PROGRAM PRG_StationProcessSettings
VAR
    bInitialised : BOOL;
    bWritePending : BOOL;
    bWriteStart : BOOL;
    bWriteBusySeen : BOOL;
    fbWritePersistentData : FB_WritePersistentData;
    stDefaultPatch : ST_PatchProcessSettings;
    stDefaultVision : ST_CameraProcessSettings;
    bSafetySaveAcceptedPending : BOOL;
    bSafetySettingsInitialised : BOOL;
    bVisionPbupSavePending : BOOL;
    bVisionPbupSaveInFlight : BOOL;
END_VAR

IF NOT bInitialised THEN
    // Preserve retained values; new speeds and delay are applied through Patch Settings.
    IF NOT ((GVL_Persistent.stPatchProcessSettings.lrDriveMotorVelocity >= 0.1) AND (GVL_Persistent.stPatchProcessSettings.lrDriveMotorVelocity <= 40)
        AND (GVL_Persistent.stPatchProcessSettings.lrPatchFeedRollVelocity >= 0.1) AND (GVL_Persistent.stPatchProcessSettings.lrPatchFeedRollVelocity <= 200)
        AND (GVL_Persistent.stPatchProcessSettings.lrWasteRollVelocity >= 0.1) AND (GVL_Persistent.stPatchProcessSettings.lrWasteRollVelocity <= 50)
        AND (GVL_Persistent.stPatchProcessSettings.udiReleaseMs >= 100) AND (GVL_Persistent.stPatchProcessSettings.udiReleaseMs <= 15000)
        AND (GVL_Persistent.stPatchProcessSettings.udiAirBlowDelayMs >= 0) AND (GVL_Persistent.stPatchProcessSettings.udiAirBlowDelayMs <= 5000)
        AND (GVL_Persistent.stPatchProcessSettings.udiDriveStopDelayMs >= 0) AND (GVL_Persistent.stPatchProcessSettings.udiDriveStopDelayMs <= 5000)) THEN
        GVL_Persistent.stPatchProcessSettings := stDefaultPatch;
        GVL_HMI.sPatchSettingsMessage := 'Stored values invalid: defaults loaded. Review and Apply.';
    ELSE
        GVL_HMI.sPatchSettingsMessage := 'Ready';
    END_IF
    GVL_HMI.stPatchProcessEdit := GVL_Persistent.stPatchProcessSettings;
    IF NOT ((GVL_Persistent.stVisionProcessSettings.udiMovingTriggerDelayMs >= 0) AND (GVL_Persistent.stVisionProcessSettings.udiMovingTriggerDelayMs <= 1000)
        AND (GVL_Persistent.stVisionProcessSettings.udiRotaryConfirmMs >= 1000) AND (GVL_Persistent.stVisionProcessSettings.udiRotaryConfirmMs <= 3000)) THEN
        GVL_Persistent.stVisionProcessSettings := stDefaultVision;
        GVL_HMI.sVisionSettingsMessage := 'Stored values invalid: defaults loaded. Review and Apply.';
    ELSE
        GVL_HMI.sVisionSettingsMessage := 'Ready';
    END_IF
    GVL_HMI.stVisionProcessEdit := GVL_Persistent.stVisionProcessSettings;
    bInitialised := TRUE;
END_IF

// Initialize the new boundary independently, including after an online source change.
IF NOT bSafetySettingsInitialised THEN
    // Reuse the existing retained door threshold; do not reset other process settings.
    IF NOT ((GVL_Config.rMainDoorHotTemperatureLimitC >= 20.0)
        AND (GVL_Config.rMainDoorHotTemperatureLimitC <= 40.0)) THEN
        GVL_Config.rMainDoorHotTemperatureLimitC := 40.0;
        GVL_HMI.sSafetySettingsMessage := 'Stored limit invalid: 40 C loaded. Review and Apply.';
    ELSE
        GVL_HMI.sSafetySettingsMessage := 'Ready';
    END_IF
    GVL_HMI.rSafetyDoorHotLimitEditC := GVL_Config.rMainDoorHotTemperatureLimitC;
    bSafetySettingsInitialised := TRUE;
END_IF

// Use existing machine status; apply before PRG_Main starts any new process.
GVL_HMI.bStationSettingsAllowed :=
    ((GVL_MASTER.stStatus.eMachineState = E_MachineState.Stopped)
     OR (GVL_MASTER.stStatus.eMachineState = E_MachineState.ReadyToStart))
    AND NOT GVL_MASTER.stStatus.stPatchDispense.bBusy
    AND NOT GVL_MASTER.stStatus.stHeatStake.bBusy
    AND NOT GVL_MASTER.stStatus.stVision.bBusy
    AND NOT GVL_Motion.stPatchFeedStatus.bBusy
    AND NOT GVL_Motion.stPatchFeedStatus.bDriveBusy
    AND NOT GVL_Motion.AxisDriveMotor.bMoving
    AND NOT GVL_Motion.AxisPatchFeedRollMotor.bMoving
    AND NOT GVL_Motion.AxisWasteRollMotor.bMoving;
bWriteStart := FALSE;

// Cancel wins over Apply. Consume command BOOLs so the HMI can issue another request.
IF GVL_HMI.bPatchSettingsCancel THEN
    GVL_HMI.stPatchProcessEdit := GVL_Persistent.stPatchProcessSettings;
    GVL_HMI.sPatchSettingsMessage := 'Edits cancelled';
ELSIF GVL_HMI.bPatchSettingsApply THEN
    IF NOT GVL_HMI.bStationSettingsAllowed THEN
        GVL_HMI.sPatchSettingsMessage := 'Apply rejected: stop machine and motion first';
    ELSIF GVL_HMI.bStationSettingsSaving THEN
        GVL_HMI.sPatchSettingsMessage := 'Apply rejected: save in progress';
    ELSIF NOT ((GVL_HMI.stPatchProcessEdit.lrDriveMotorVelocity >= 0.1) AND (GVL_HMI.stPatchProcessEdit.lrDriveMotorVelocity <= 40)
        AND (GVL_HMI.stPatchProcessEdit.lrPatchFeedRollVelocity >= 0.1) AND (GVL_HMI.stPatchProcessEdit.lrPatchFeedRollVelocity <= 200)
        AND (GVL_HMI.stPatchProcessEdit.lrWasteRollVelocity >= 0.1) AND (GVL_HMI.stPatchProcessEdit.lrWasteRollVelocity <= 50)
        AND (GVL_HMI.stPatchProcessEdit.udiReleaseMs >= 100) AND (GVL_HMI.stPatchProcessEdit.udiReleaseMs <= 15000)
        AND (GVL_HMI.stPatchProcessEdit.udiAirBlowDelayMs >= 0) AND (GVL_HMI.stPatchProcessEdit.udiAirBlowDelayMs <= 5000)
        AND (GVL_HMI.stPatchProcessEdit.udiDriveStopDelayMs >= 0) AND (GVL_HMI.stPatchProcessEdit.udiDriveStopDelayMs <= 5000)) THEN
        GVL_HMI.sPatchSettingsMessage := 'Apply rejected: value outside allowed range';
    ELSE
        GVL_Persistent.stPatchProcessSettings := GVL_HMI.stPatchProcessEdit;
        bWritePending := TRUE;
        GVL_HMI.bStationSettingsSaveError := FALSE;
        GVL_HMI.udiStationSettingsSaveErrorId := 0;
        GVL_HMI.sPatchSettingsMessage := 'Applied - saving';
    END_IF
END_IF
GVL_HMI.bPatchSettingsApply := FALSE;
GVL_HMI.bPatchSettingsCancel := FALSE;
GVL_HMI.stPatchProcessApplied := GVL_Persistent.stPatchProcessSettings;

// Cancel wins over Apply. Consume command BOOLs so the HMI can issue another request.
IF GVL_HMI.bVisionSettingsCancel THEN
    GVL_HMI.stVisionProcessEdit := GVL_Persistent.stVisionProcessSettings;
    GVL_HMI.sVisionSettingsMessage := 'Edits cancelled';
ELSIF GVL_HMI.bVisionSettingsApply THEN
    IF NOT GVL_HMI.bStationSettingsAllowed THEN
        GVL_HMI.sVisionSettingsMessage := 'Apply rejected: stop machine and motion first';
    ELSIF GVL_HMI.bStationSettingsSaving THEN
        GVL_HMI.sVisionSettingsMessage := 'Apply rejected: save in progress';
    ELSIF NOT ((GVL_HMI.stVisionProcessEdit.udiMovingTriggerDelayMs >= 0) AND (GVL_HMI.stVisionProcessEdit.udiMovingTriggerDelayMs <= 1000)
        AND (GVL_HMI.stVisionProcessEdit.udiRotaryConfirmMs >= 1000) AND (GVL_HMI.stVisionProcessEdit.udiRotaryConfirmMs <= 3000)) THEN
        GVL_HMI.sVisionSettingsMessage := 'Apply rejected: value outside allowed range';
    ELSE
        GVL_Persistent.stVisionProcessSettings := GVL_HMI.stVisionProcessEdit;
        bWritePending := TRUE;
        GVL_HMI.bStationSettingsSaveError := FALSE;
        GVL_HMI.udiStationSettingsSaveErrorId := 0;
        GVL_HMI.sVisionSettingsMessage := 'Applied - saving';
    END_IF
END_IF
GVL_HMI.bVisionSettingsApply := FALSE;
GVL_HMI.bVisionSettingsCancel := FALSE;
GVL_HMI.stVisionProcessApplied := GVL_Persistent.stVisionProcessSettings;

// Safety settings are accepted only while Stopped and all existing settings/motion gates are clear.
GVL_HMI.bSafetySettingsAllowed := GVL_HMI.bStationSettingsAllowed
    AND (GVL_MASTER.stStatus.eMachineState = E_MachineState.Stopped)
    AND NOT GVL_MASTER.stCommand.bReset;
IF GVL_HMI.bSafetySettingsCancel THEN
    GVL_HMI.rSafetyDoorHotLimitEditC := GVL_Config.rMainDoorHotTemperatureLimitC;
    GVL_HMI.sSafetySettingsMessage := 'Edits cancelled';
ELSIF GVL_HMI.bSafetySettingsApply THEN
    IF NOT GVL_HMI.bSafetySettingsAllowed THEN
        GVL_HMI.sSafetySettingsMessage := 'Apply rejected: machine must be Stopped and idle';
    ELSIF GVL_HMI.bStationSettingsSaving THEN
        GVL_HMI.sSafetySettingsMessage := 'Apply rejected: save in progress';
    ELSIF NOT ((GVL_HMI.rSafetyDoorHotLimitEditC >= 20.0)
        AND (GVL_HMI.rSafetyDoorHotLimitEditC <= 40.0)) THEN
        GVL_HMI.sSafetySettingsMessage := 'Apply rejected: allowed range 20 to 40 C';
    ELSE
        GVL_Config.rMainDoorHotTemperatureLimitC := GVL_HMI.rSafetyDoorHotLimitEditC;
        bWritePending := TRUE;
        bSafetySaveAcceptedPending := TRUE;
        GVL_HMI.bStationSettingsSaveError := FALSE;
        GVL_HMI.udiStationSettingsSaveErrorId := 0;
        GVL_HMI.sSafetySettingsMessage := 'Applied - saving';
    END_IF
END_IF
GVL_HMI.bSafetySettingsApply := FALSE;
GVL_HMI.bSafetySettingsCancel := FALSE;
GVL_HMI.rSafetyDoorHotLimitAppliedC := GVL_Config.rMainDoorHotTemperatureLimitC;

// Request is latched by PRG_Main after this program; consume it on the next scan.
IF GVL_HMI.bVisionPbupSaveRequest THEN
    GVL_HMI.bVisionPbupSaveRequest := FALSE;
    bWritePending := TRUE;
    bVisionPbupSavePending := TRUE;
    GVL_HMI.bVisionPbupSaveError := FALSE;
    GVL_HMI.udiVisionPbupSaveErrorId := 0;
    GVL_HMI.sVisionPbupSaveStatus := 'PBUP state: save pending';
END_IF
IF bWritePending AND NOT fbWritePersistentData.BUSY THEN
    bWriteStart := TRUE;
    bWritePending := FALSE;
    bWriteBusySeen := FALSE;
END_IF
IF bWriteStart AND bVisionPbupSavePending THEN
    bVisionPbupSavePending := FALSE;
    bVisionPbupSaveInFlight := TRUE;
    GVL_HMI.sVisionPbupSaveStatus := 'PBUP state: saving';
END_IF
fbWritePersistentData(NETID := '', PORT := 851, START := bWriteStart,
    TMOUT := T#2S, MODE := SPDM_VAR_BOOST);
IF fbWritePersistentData.BUSY THEN bWriteBusySeen := TRUE; END_IF
IF fbWritePersistentData.ERR THEN
    IF bVisionPbupSaveInFlight THEN
        bVisionPbupSaveInFlight := FALSE;
        GVL_HMI.bVisionPbupSaveError := TRUE;
        GVL_HMI.udiVisionPbupSaveErrorId := fbWritePersistentData.ERRID;
        GVL_HMI.sVisionPbupSaveStatus := 'PBUP state: SAVE FAILED; confirm state again to retry';
    END_IF
    GVL_HMI.bStationSettingsSaveError := TRUE;
    GVL_HMI.udiStationSettingsSaveErrorId := fbWritePersistentData.ERRID;
    IF bSafetySaveAcceptedPending THEN
        GVL_HMI.sSafetySettingsMessage := 'Applied, SAVE FAILED. Correct cause and Apply again.';
        bSafetySaveAcceptedPending := FALSE;
    END_IF
    IF GVL_HMI.sPatchSettingsMessage = 'Applied - saving' THEN
        GVL_HMI.sPatchSettingsMessage := 'Applied, SAVE FAILED. Correct cause and Apply again.';
    END_IF
    IF GVL_HMI.sVisionSettingsMessage = 'Applied - saving' THEN
        GVL_HMI.sVisionSettingsMessage := 'Applied, SAVE FAILED. Correct cause and Apply again.';
    END_IF
ELSIF bWriteBusySeen AND NOT fbWritePersistentData.BUSY THEN
    IF bVisionPbupSaveInFlight THEN
        bVisionPbupSaveInFlight := FALSE;
        GVL_HMI.sVisionPbupSaveStatus := 'PBUP state: saved';
    END_IF
    bWriteBusySeen := FALSE;
    IF bSafetySaveAcceptedPending THEN
        GVL_HMI.sSafetySettingsMessage := 'Applied and saved';
        bSafetySaveAcceptedPending := FALSE;
    END_IF
    IF GVL_HMI.sPatchSettingsMessage = 'Applied - saving' THEN
        GVL_HMI.sPatchSettingsMessage := 'Applied and saved';
    END_IF
    IF GVL_HMI.sVisionSettingsMessage = 'Applied - saving' THEN
        GVL_HMI.sVisionSettingsMessage := 'Applied and saved';
    END_IF
END_IF
GVL_HMI.bStationSettingsSaving := fbWritePersistentData.BUSY OR bWritePending OR bWriteStart;
// Preserve direction, NC dynamics, watchdogs and temporary feedback configuration.
GVL_Motion.stPatchFeedSettings.lrDriveMotorVelocity := GVL_Persistent.stPatchProcessSettings.lrDriveMotorVelocity;
GVL_Motion.stPatchFeedSettings.lrPatchFeedRollVelocity := GVL_Persistent.stPatchProcessSettings.lrPatchFeedRollVelocity;
GVL_Motion.stPatchFeedSettings.lrWasteRollVelocity := GVL_Persistent.stPatchProcessSettings.lrWasteRollVelocity;

// Patch vertical sensors are fitted: physical feedback is mandatory, including after an online change.
GVL_Motion.stPatchFeedSettings.bUsePatchVerticalFeedback := TRUE;

GVL_HMI.bVisionPbupSaving := bVisionPbupSavePending OR bVisionPbupSaveInFlight
    OR GVL_HMI.bVisionPbupSaveRequest;

END_PROGRAM

(* stored: Version 1.1.0.1, ProductVersion 3.1.4026.18
   POU PRG_StationProcessSettings: Id {3e164b6f-de11-4dca-9030-f5df8bd57159}, SpecialFunc None *)
